// TIA Portal V20 export
// export: Created 2026-10-12T16:46:22.3324652Z, ExportSetting WithDefaults, DisplayName Totally Integrated Automation Portal, DisplayVersion V20 Update 6, DisplayName TIA Portal Openness, DisplayVersion V20 Update 6, DisplayName TIA Portal Version Control Interface, DisplayVersion V20 Update 6, DisplayName SINAMICS Startdrive Advanced, DisplayVersion V20 SP1 Update 2, DisplayName SINAMICS Startdrive G110M, G120, G120C, G120D, G120P, G115D, DisplayVersion V20 SP1 Update 2, DisplayName SINAMICS Startdrive G130, G150, S120, S150, SINAMICS MV, G220, S200, S210, DisplayVersion V20 SP1 Update 2, DisplayName STEP 7 Professional, DisplayVersion V20 Update 6, DisplayName STEP 7 Safety, DisplayVersion V20 Update 2, DisplayName WinCC Basic/Comfort/Advanced, DisplayVersion V20 Update 6, DisplayName WinCC Professional, DisplayVersion V20 Update 6, DisplayName WinCC Unified, DisplayVersion V20 Update 6
VAR_GLOBAL   // PLC tag table "KP8_Neu"
   KP8_1_IB_Tasten AT %IB1000 : Byte;   // IB_Tasten
   KP8_1_IB_DI AT %IB1001 : Byte;   // IB_DI
   KP8_2_IB_Tasten AT %IB2000 : Byte;   // IB_Tasten
   KP8_2_IB_DI AT %IB2001 : Byte;   // IB_DI
   KP8_3_IB_Tasten AT %IB3000 : Byte;   // IB_Tasten
   KP8_3_IB_DI AT %IB3001 : Byte;   // IB_DI
   KP8_4_IB_Tasten AT %IB4000 : Byte;   // IB_Tasten
   KP8_4_IB_DI AT %IB4001 : Byte;   // IB_DI
   KP8_5_IB_Tasten AT %IB5000 : Byte;   // IB_Tasten
   KP8_5_IB_DI AT %IB5001 : Byte;   // IB_DI
   KP8_6_IB_Tasten AT %IB6000 : Byte;   // IB_Tasten
   KP8_6_IB_DI AT %IB6001 : Byte;   // IB_DI
   KP8_7_IB_Tasten AT %IB7000 : Byte;   // IB_Tasten
   KP8_7_IB_DI AT %IB7001 : Byte;   // IB_DI
   KP8_8_IB_Tasten AT %IB8000 : Byte;   // IB_Tasten
   KP8_8_IB_DI AT %IB8001 : Byte;   // IB_DI
   KP8_9_IB_Tasten AT %IB9000 : Byte;   // IB_Tasten
   KP8_9_IB_DI AT %IB9001 : Byte;   // IB_DI
   KP8_10_IB_Tasten AT %IB10000 : Byte;   // IB_Tasten
   KP8_10_IB_DI AT %IB10001 : Byte;   // IB_DI
   KP8_11_IB_Tasten AT %IB11000 : Byte;   // IB_Tasten
   KP8_11_IB_DI AT %IB11001 : Byte;   // IB_DI
   KP8_12_IB_Tasten AT %IB12000 : Byte;   // IB_Tasten
   KP8_12_IB_DI AT %IB12001 : Byte;   // IB_DI
   KP8_13_IB_Tasten AT %IB13000 : Byte;   // IB_Tasten
   KP8_13_IB_DI AT %IB13001 : Byte;   // IB_DI
   KP8_14_IB_Tasten AT %IB14000 : Byte;   // IB_Tasten
   KP8_14_IB_DI AT %IB14001 : Byte;   // IB_DI
   KP8_15_IB_Tasten AT %IB15000 : Byte;   // IB_Tasten
   KP8_15_IB_DI AT %IB15001 : Byte;   // IB_DI
   KP8_16_IB_Tasten AT %IB16000 : Byte;   // IB_Tasten
   KP8_16_IB_DI AT %IB16001 : Byte;   // IB_DI
   KP8_17_IB_Tasten AT %IB17000 : Byte;   // IB_Tasten
   KP8_17_IB_DI AT %IB17001 : Byte;   // IB_DI
   KP8_18_IB_Tasten AT %IB18000 : Byte;   // IB_Tasten
   KP8_18_IB_DI AT %IB18001 : Byte;   // IB_DI
   KP8_19_IB_Tasten AT %IB19000 : Byte;   // IB_Tasten
   KP8_19_IB_DI AT %IB19001 : Byte;   // IB_DI
   KP8_20_IB_Tasten AT %IB20000 : Byte;   // IB_Tasten
   KP8_20_IB_DI AT %IB20001 : Byte;   // IB_DI
   KP8_21_IB_Tasten AT %IB21000 : Byte;   // IB_Tasten
   KP8_21_IB_DI AT %IB21001 : Byte;   // IB_DI
   KP8_22_IB_Tasten AT %IB22000 : Byte;   // IB_Tasten
   KP8_22_IB_DI AT %IB22001 : Byte;   // IB_DI
   KP8_23_IB_Tasten AT %IB23000 : Byte;   // IB_Tasten
   KP8_23_IB_DI AT %IB23001 : Byte;   // IB_DI
   KP8_24_IB_Tasten AT %IB24000 : Byte;   // IB_Tasten
   KP8_24_IB_DI AT %IB24001 : Byte;   // IB_DI
   KP8_25_IB_Tasten AT %IB25000 : Byte;   // IB_Tasten
   KP8_25_IB_DI AT %IB25001 : Byte;   // IB_DI
   KP8_26_IB_Tasten AT %IB26000 : Byte;   // IB_Tasten
   KP8_26_IB_DI AT %IB26001 : Byte;   // IB_DI
   KP8_27_IB_Tasten AT %IB27000 : Byte;   // IB_Tasten
   KP8_27_IB_DI AT %IB27001 : Byte;   // IB_DI
   KP8_28_IB_Tasten AT %IB28000 : Byte;   // IB_Tasten
   KP8_28_IB_DI AT %IB28001 : Byte;   // IB_DI
   KP8_1_QB_Rot AT %QB1000 : Byte;   // QB_Rot
   KP8_1_QB_Gruen AT %QB1001 : Byte;   // QB_Gruen
   KP8_1_QB_Blau AT %QB1002 : Byte;   // QB_Blau
   KP8_1_QB_DO AT %QB1003 : Byte;   // QB_DO
   KP8_2_QB_Rot AT %QB2000 : Byte;   // QB_Rot
   KP8_2_QB_Gruen AT %QB2001 : Byte;   // QB_Gruen
   KP8_2_QB_Blau AT %QB2002 : Byte;   // QB_Blau
   KP8_2_QB_DO AT %QB2003 : Byte;   // QB_DO
   KP8_3_QB_Rot AT %QB3000 : Byte;   // QB_Rot
   KP8_3_QB_Gruen AT %QB3001 : Byte;   // QB_Gruen
   KP8_3_QB_Blau AT %QB3002 : Byte;   // QB_Blau
   KP8_3_QB_DO AT %QB3003 : Byte;   // QB_DO
   KP8_4_QB_Rot AT %QB4000 : Byte;   // QB_Rot
   KP8_4_QB_Gruen AT %QB4001 : Byte;   // QB_Gruen
   KP8_4_QB_Blau AT %QB4002 : Byte;   // QB_Blau
   KP8_4_QB_DO AT %QB4003 : Byte;   // QB_DO
   KP8_5_QB_Rot AT %QB5000 : Byte;   // QB_Rot
   KP8_5_QB_Gruen AT %QB5001 : Byte;   // QB_Gruen
   KP8_5_QB_Blau AT %QB5002 : Byte;   // QB_Blau
   KP8_5_QB_DO AT %QB5003 : Byte;   // QB_DO
   KP8_6_QB_Rot AT %QB6000 : Byte;   // QB_Rot
   KP8_6_QB_Gruen AT %QB6001 : Byte;   // QB_Gruen
   KP8_6_QB_Blau AT %QB6002 : Byte;   // QB_Blau
   KP8_6_QB_DO AT %QB6003 : Byte;   // QB_DO
   KP8_7_QB_Rot AT %QB7000 : Byte;   // QB_Rot
   KP8_7_QB_Gruen AT %QB7001 : Byte;   // QB_Gruen
   KP8_7_QB_Blau AT %QB7002 : Byte;   // QB_Blau
   KP8_7_QB_DO AT %QB7003 : Byte;   // QB_DO
   KP8_8_QB_Rot AT %QB8000 : Byte;   // QB_Rot
   KP8_8_QB_Gruen AT %QB8001 : Byte;   // QB_Gruen
   KP8_8_QB_Blau AT %QB8002 : Byte;   // QB_Blau
   KP8_8_QB_DO AT %QB8003 : Byte;   // QB_DO
   KP8_9_QB_Rot AT %QB9000 : Byte;   // QB_Rot
   KP8_9_QB_Gruen AT %QB9001 : Byte;   // QB_Gruen
   KP8_9_QB_Blau AT %QB9002 : Byte;   // QB_Blau
   KP8_9_QB_DO AT %QB9003 : Byte;   // QB_DO
   KP8_10_QB_Rot AT %QB10000 : Byte;   // QB_Rot
   KP8_10_QB_Gruen AT %QB10001 : Byte;   // QB_Gruen
   KP8_10_QB_Blau AT %QB10002 : Byte;   // QB_Blau
   KP8_10_QB_DO AT %QB10003 : Byte;   // QB_DO
   KP8_11_QB_Rot AT %QB11000 : Byte;   // QB_Rot
   KP8_11_QB_Gruen AT %QB11001 : Byte;   // QB_Gruen
   KP8_11_QB_Blau AT %QB11002 : Byte;   // QB_Blau
   KP8_11_QB_DO AT %QB11003 : Byte;   // QB_DO
   KP8_12_QB_Rot AT %QB12000 : Byte;   // QB_Rot
   KP8_12_QB_Gruen AT %QB12001 : Byte;   // QB_Gruen
   KP8_12_QB_Blau AT %QB12002 : Byte;   // QB_Blau
   KP8_12_QB_DO AT %QB12003 : Byte;   // QB_DO
   KP8_13_QB_Rot AT %QB13000 : Byte;   // QB_Rot
   KP8_13_QB_Gruen AT %QB13001 : Byte;   // QB_Gruen
   KP8_13_QB_Blau AT %QB13002 : Byte;   // QB_Blau
   KP8_13_QB_DO AT %QB13003 : Byte;   // QB_DO
   KP8_14_QB_Rot AT %QB14000 : Byte;   // QB_Rot
   KP8_14_QB_Gruen AT %QB14001 : Byte;   // QB_Gruen
   KP8_14_QB_Blau AT %QB14002 : Byte;   // QB_Blau
   KP8_14_QB_DO AT %QB14003 : Byte;   // QB_DO
   KP8_15_QB_Rot AT %QB15000 : Byte;   // QB_Rot
   KP8_15_QB_Gruen AT %QB15001 : Byte;   // QB_Gruen
   KP8_15_QB_Blau AT %QB15002 : Byte;   // QB_Blau
   KP8_15_QB_DO AT %QB15003 : Byte;   // QB_DO
   KP8_16_QB_Rot AT %QB16000 : Byte;   // QB_Rot
   KP8_16_QB_Gruen AT %QB16001 : Byte;   // QB_Gruen
   KP8_16_QB_Blau AT %QB16002 : Byte;   // QB_Blau
   KP8_16_QB_DO AT %QB16003 : Byte;   // QB_DO
   KP8_17_QB_Rot AT %QB17000 : Byte;   // QB_Rot
   KP8_17_QB_Gruen AT %QB17001 : Byte;   // QB_Gruen
   KP8_17_QB_Blau AT %QB17002 : Byte;   // QB_Blau
   KP8_17_QB_DO AT %QB17003 : Byte;   // QB_DO
   KP8_18_QB_Rot AT %QB18000 : Byte;   // QB_Rot
   KP8_18_QB_Gruen AT %QB18001 : Byte;   // QB_Gruen
   KP8_18_QB_Blau AT %QB18002 : Byte;   // QB_Blau
   KP8_18_QB_DO AT %QB18003 : Byte;   // QB_DO
   KP8_19_QB_Rot AT %QB19000 : Byte;   // QB_Rot
   KP8_19_QB_Gruen AT %QB19001 : Byte;   // QB_Gruen
   KP8_19_QB_Blau AT %QB19002 : Byte;   // QB_Blau
   KP8_19_QB_DO AT %QB19003 : Byte;   // QB_DO
   KP8_20_QB_Rot AT %QB20000 : Byte;   // QB_Rot
   KP8_20_QB_Gruen AT %QB20001 : Byte;   // QB_Gruen
   KP8_20_QB_Blau AT %QB20002 : Byte;   // QB_Blau
   KP8_20_QB_DO AT %QB20003 : Byte;   // QB_DO
   KP8_21_QB_Rot AT %QB21000 : Byte;   // QB_Rot
   KP8_21_QB_Gruen AT %QB21001 : Byte;   // QB_Gruen
   KP8_21_QB_Blau AT %QB21002 : Byte;   // QB_Blau
   KP8_21_QB_DO AT %QB21003 : Byte;   // QB_DO
   KP8_22_QB_Rot AT %QB22000 : Byte;   // QB_Rot
   KP8_22_QB_Gruen AT %QB22001 : Byte;   // QB_Gruen
   KP8_22_QB_Blau AT %QB22002 : Byte;   // QB_Blau
   KP8_22_QB_DO AT %QB22003 : Byte;   // QB_DO
   KP8_23_QB_Rot AT %QB23000 : Byte;   // QB_Rot
   KP8_23_QB_Gruen AT %QB23001 : Byte;   // QB_Gruen
   KP8_23_QB_Blau AT %QB23002 : Byte;   // QB_Blau
   KP8_23_QB_DO AT %QB23003 : Byte;   // QB_DO
   KP8_24_QB_Rot AT %QB24000 : Byte;   // QB_Rot
   KP8_24_QB_Gruen AT %QB24001 : Byte;   // QB_Gruen
   KP8_24_QB_Blau AT %QB24002 : Byte;   // QB_Blau
   KP8_24_QB_DO AT %QB24003 : Byte;   // QB_DO
   KP8_25_QB_Rot AT %QB25000 : Byte;   // QB_Rot
   KP8_25_QB_Gruen AT %QB25001 : Byte;   // QB_Gruen
   KP8_25_QB_Blau AT %QB25002 : Byte;   // QB_Blau
   KP8_25_QB_DO AT %QB25003 : Byte;   // QB_DO
   KP8_26_QB_Rot AT %QB26000 : Byte;   // QB_Rot
   KP8_26_QB_Gruen AT %QB26001 : Byte;   // QB_Gruen
   KP8_26_QB_Blau AT %QB26002 : Byte;   // QB_Blau
   KP8_26_QB_DO AT %QB26003 : Byte;   // QB_DO
   KP8_27_QB_Rot AT %QB27000 : Byte;   // QB_Rot
   KP8_27_QB_Gruen AT %QB27001 : Byte;   // QB_Gruen
   KP8_27_QB_Blau AT %QB27002 : Byte;   // QB_Blau
   KP8_27_QB_DO AT %QB27003 : Byte;   // QB_DO
   KP8_28_QB_Rot AT %QB28000 : Byte;   // QB_Rot
   KP8_28_QB_Gruen AT %QB28001 : Byte;   // QB_Gruen
   KP8_28_QB_Blau AT %QB28002 : Byte;   // QB_Blau
   KP8_28_QB_DO AT %QB28003 : Byte;   // QB_DO
END_VAR
